# EPICS substitutions: b-55B2VNC/src/main/epics/PCF0CoreApp/Db/StateMachine.substitutions
file "nds3_StateMachine.template"{
pattern
{
    BOARDTYPE,
    BOARDTYPEIDX,
    CBS1,
    CBS2,
    STATEMACHINE_PARENT,
    STATEMACHINE_NAME
}
{
    "B",
    "0",
    "TEST",
    "FCT0",
    "",
    "StateMachine"
}
}
file "nds3_StateMachine.template"{
pattern
{
    BOARDTYPE,
    BOARDTYPEIDX,
    CBS1,
    CBS2,
    STATEMACHINE_PARENT,
    STATEMACHINE_NAME
}
{
    "B",
    "8",
    "D1",
    "I2",
    "",
    "StateMachine"
}
}
